Staubli VAL3: Force4Item.pjx

--- Force4Item.pjx ---
Parameters version=s8.15.3Cs9_BS3337 stackSize=5000 millimeterUnit=true
Program file=start.pgx
Program file=stop.pgx
Data file=Force4Item.dtx

--- Force4Item.dtx ---
mdesc mNomSpeed
public string sArmType
public num nMaxJnt4Force[4]

--- start.pgx ---
program start()
begin
end

--- stop.pgx ---
program stop()
begin
end
